Fanuc KAREL source: ko00041.KL

-- PROVISIONAL review KL for V770-1; original PC SHA256 486ec2265fe29498fcdda0df1ef52f390ff49c0469c900f2fd5722d6fbbd2cf6
-- Incomplete behavior may be omitted. Consult companion uncertainty JSON. Do not deploy.
PROGRAM KO00041
%NOLOCKGROUP
BEGIN
  -- UNRESOLVED_PC offsets 5-12; opcodes 9D,23
  -- UNRESOLVED_PC offsets 17-69; opcodes 27,27,49,7E,AD,27,49,7E,AD,22,31,7E,4A
  -- UNRESOLVED_PC offsets 74-78; opcodes 7F
END KO00041
